Fanuc KAREL source: kd00047.KL

-- PROVISIONAL review KL for V940-1; original PC SHA256 348f76738a9ebfd8d93a47e68de620e40bb07c5dc43f8ff35c8cdb1a5d54a96e
-- Incomplete behavior may be omitted. Consult companion uncertainty JSON. Do not deploy.
PROGRAM KD00047
%NOLOCKGROUP
VAR
  I : INTEGER
  J : INTEGER
  B : BOOLEAN
  R : REAL
  S : STRING[80]
-- UNRESOLVED_DECL V type=000013
BEGIN
  -- V9_ZERO_TABLE_METADATA_HINT layout=0001; no indexed target words; source/name/runtime held
  -- UNRESOLVED_PC offsets 5-20; opcodes 2E,22,32,35
  -- UNRESOLVED_PC offsets 25-46; opcodes 01,49,2E,0A,82,0B
  -- UNRESOLVED_PC offsets 51-55; opcodes 7F
END KD00047
